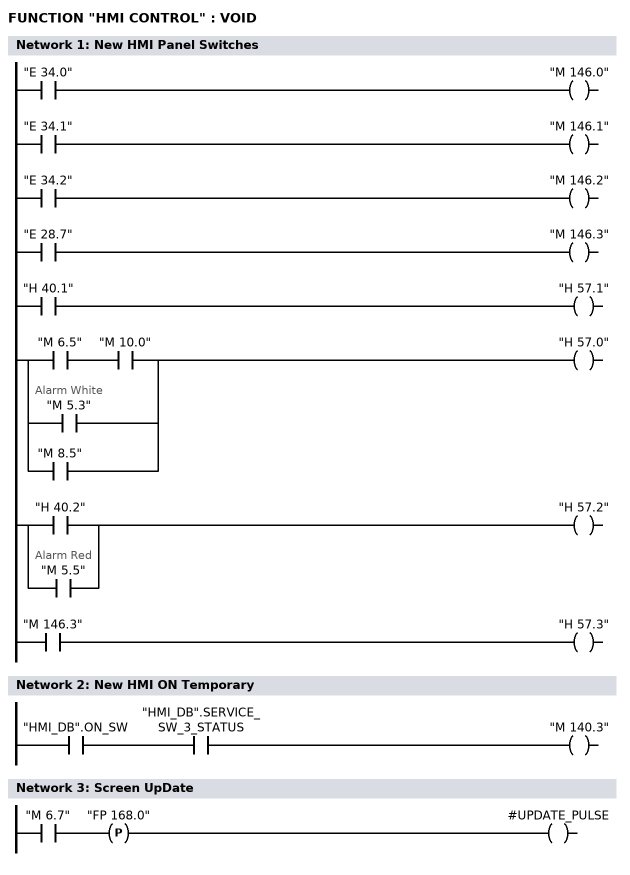

      A     "E 34.0";
      =     "M 146.0";
//;
      A     "E 34.1";
      =     "M 146.1";
//;
      A     "E 34.2";
      =     "M 146.2";
//;
      A     "E 28.7";
      =     "M 146.3";
//;
      A     "H 40.1";
      =     "H 57.1";
//;
      A(    ;
      A     "M 6.5";
      A     "M 10.0";
      )     ;
      O     "M 5.3"; // Alarm White
      O     "M 8.5";
      =     "H 57.0";
//;
      A     "H 40.2";
      O     "M 5.5"; // Alarm Red
      =     "H 57.2";
//;
      A     "M 146.3";
      =     "H 57.3";
NETWORK
TITLE =New HMI ON Temporary

      A     "HMI_DB".ON_SW;
      A     "HMI_DB".SERVICE_SW_3_STATUS;
      =     "M 140.3";
NETWORK
TITLE =Screen UpDate

      A     "M 6.7";
      FP    "FP 168.0";
      =     #UPDATE_PULSE;
NETWORK
TITLE =Screen 0 Soft Switches

      A(    ;
      L     "HMI_DB".ACTUAL_HMI_SCREEN_NO;
      L     "HMI_UPDATE".HMI_MAIN_PAGE_GRAPHIC;
      <>I   ;
      )     ;
      O     #UPDATE_PULSE;
      JNB   MAIN;
NETWORK
TITLE =Service Switch Status - Screen 0 SSW Inputs
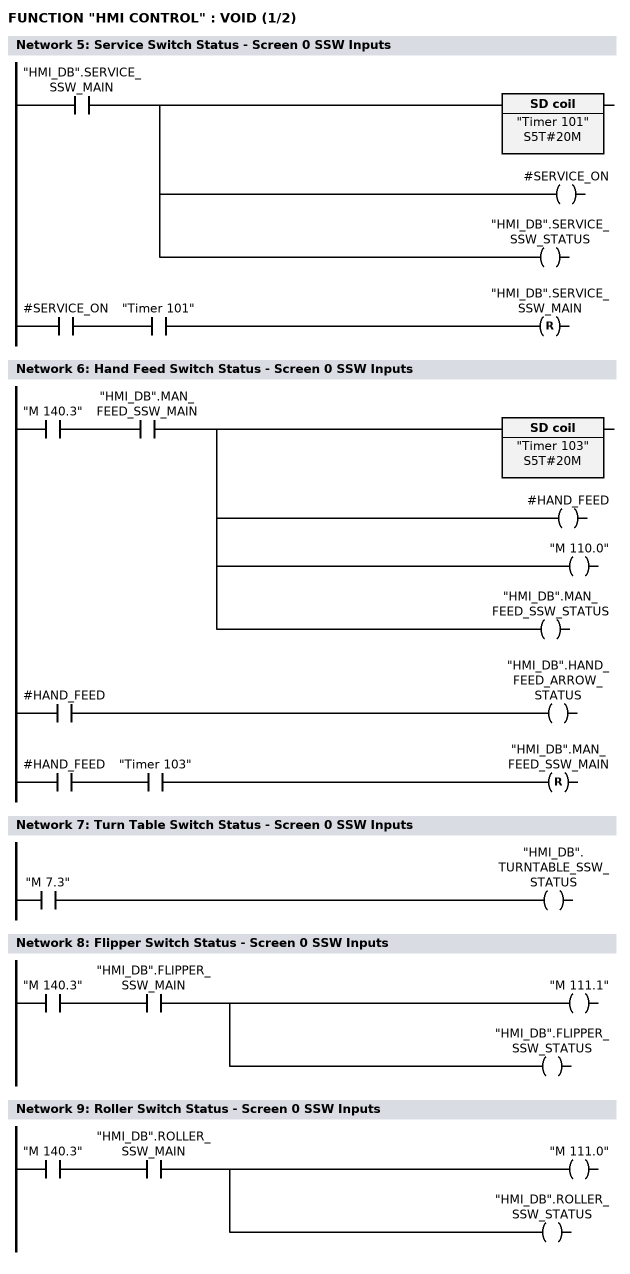

      A     "HMI_DB".SERVICE_SSW_MAIN;
      L     S5T#20M;
      SD    "Timer 101";
      =     #SERVICE_ON;
      =     "HMI_DB".SERVICE_SSW_STATUS;
//;
      A     #SERVICE_ON;
      A     "Timer 101";
      R     "HMI_DB".SERVICE_SSW_MAIN;
NETWORK
TITLE =Hand Feed Switch Status - Screen 0 SSW Inputs

      A     "M 140.3";
      A     "HMI_DB".MAN_FEED_SSW_MAIN;
      L     S5T#20M;
      SD    "Timer 103";
      =     #HAND_FEED;
      =     "M 110.0";
      =     "HMI_DB".MAN_FEED_SSW_STATUS;
//;
      A     #HAND_FEED;
      =     "HMI_DB".HAND_FEED_ARROW_STATUS;
//;
      A     #HAND_FEED;
      A     "Timer 103";
      R     "HMI_DB".MAN_FEED_SSW_MAIN;
NETWORK
TITLE =Turn Table Switch Status - Screen 0 SSW Inputs

      A     "M 7.3";
      =     "HMI_DB".TURNTABLE_SSW_STATUS;
NETWORK
TITLE =Flipper Switch Status - Screen 0 SSW Inputs

      A     "M 140.3";
      A     "HMI_DB".FLIPPER_SSW_MAIN;
      =     "M 111.1";
      =     "HMI_DB".FLIPPER_SSW_STATUS;
NETWORK
TITLE =Roller Switch Status - Screen 0 SSW Inputs

      A     "M 140.3";
      A     "HMI_DB".ROLLER_SSW_MAIN;
      =     "M 111.0";
      =     "HMI_DB".ROLLER_SSW_STATUS;
NETWORK
TITLE =HMI Service Switch Reset
//HMI Service Switch Reset when 2145 Exits Packets + 10s Delay
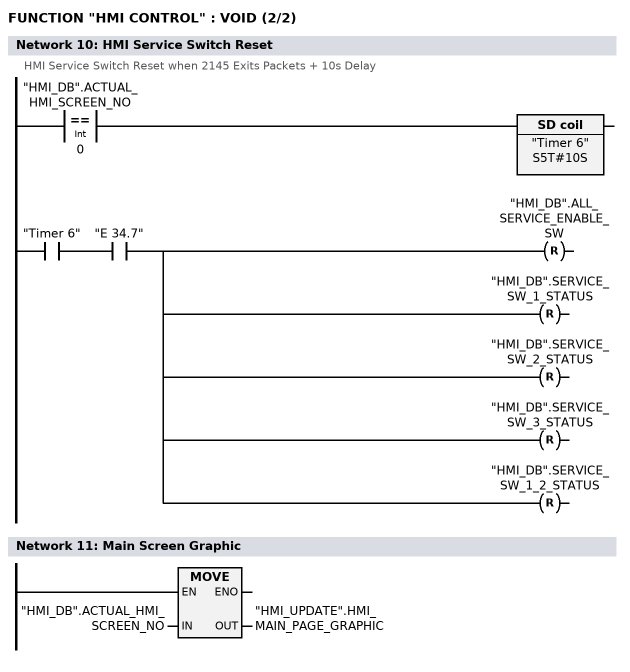
      A(    ;
      L     "HMI_DB".ACTUAL_HMI_SCREEN_NO;
      L     0;
      ==I   ;
      )     ;
      L     S5T#10S;
      SD    "Timer 6";
//;
      A     "Timer 6";
      A     "E 34.7";
      R     "HMI_DB".ALL_SERVICE_ENABLE_SW;
      R     "HMI_DB".SERVICE_SW_1_STATUS;
      R     "HMI_DB".SERVICE_SW_2_STATUS;
      R     "HMI_DB".SERVICE_SW_3_STATUS;
      R     "HMI_DB".SERVICE_SW_1_2_STATUS;
NETWORK
TITLE =Main Screen Graphic


      L     "HMI_DB".ACTUAL_HMI_SCREEN_NO;
      T     "HMI_UPDATE".HMI_MAIN_PAGE_GRAPHIC;

MAIN: NOP   0;
END_FUNCTION

FUNCTION "HMI COMMS" : VOID
TITLE =HMI Communications
//OMRON NS12  on DB12
NAME : HMI_COMM
VERSION : 0.1


VAR_TEMP
  UPDATE_PULSE_0 : BOOL ;
  UPDATE_PULSE_1 : BOOL ;
  UPDATE_PULSE_2 : BOOL ;
  UPDATE_PULSE_3 : BOOL ;
  UPDATE_PULSE_4 : BOOL ;
  UPDATE_PULSE_5 : BOOL ;
  UPDATE_PULSE_6 : BOOL ;
  UPDATE_1 : BOOL ;
  UPDATE_2 : BOOL ;
  UPDATE_3 : BOOL ;
  UPDATE_4 : BOOL ;
  UPDATE_5 : BOOL ;
  UPDATE_6 : BOOL ;
  UPDATE_7 : BOOL ;
  UPDATE_8 : BOOL ;
  UPDATE_9 : BOOL ;
  UPDATE_10 : BOOL ;
  UPDATE_11 : BOOL ;
  UPDATE_12 : BOOL ;
  UPDATE_13 : BOOL ;
  TEMP1 : BOOL ;
  TEST : BOOL ;
  CONVEYOR_0_COLOR : BYTE ;
  ELEVATOR_COLOR : BYTE ;
  CONVEYOR_1_COLOR : BYTE ;
  CONVEYOR_2_COLOR : BYTE ;
  CONVEYOR_3_COLOR : BYTE ;
  CONVEYOR_4_COLOR : BYTE ;
  CONVEYOR_5_COLOR : BYTE ;
  CONVEYOR_6_COLOR : BYTE ;
  CONVEYOR_7_COLOR : BYTE ;
  CONVEYOR_8_COLOR : BYTE ;
  CONVEYOR_9_COLOR : BYTE ;
  PUSHER_2_COLOR : BOOL ;
  CONVEYOR_11_COLOR : BYTE ;
  CONVEYOR_12_COLOR : BYTE ;
  CONVEYOR_13_COLOR : BYTE ;
  CONVEYOR_21_COLOR : BYTE ;
  CONVEYOR_22_COLOR : BYTE ;
  CONVEYOR_23_COLOR : BYTE ;
  CONVEYOR_10_COLOR : BYTE ;
  NEW_ORDER_COLOR : BYTE ;
END_VAR
BEGIN
NETWORK
TITLE =HMI - UpDate Timing
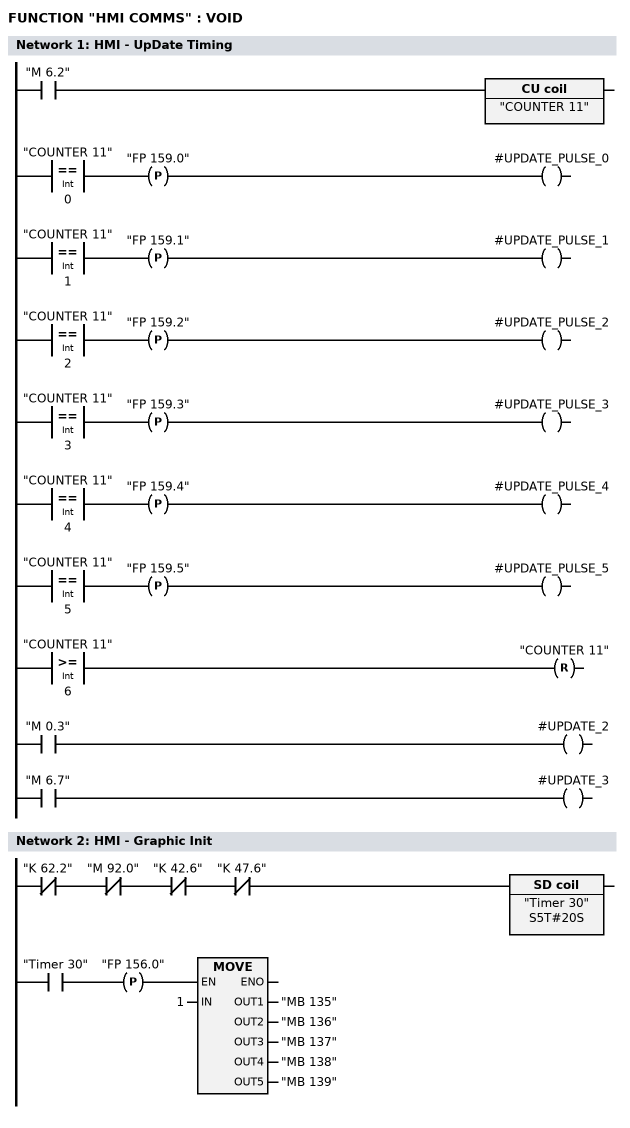

      A     "M 6.2";
      CU    "COUNTER 11";
//;
      A(    ;
      L     "COUNTER 11";
      L     0;
      ==I   ;
      )     ;
      FP    "FP 159.0";
      =     #UPDATE_PULSE_0;
//;
      A(    ;
      L     "COUNTER 11";
      L     1;
      ==I   ;
      )     ;
      FP    "FP 159.1";
      =     #UPDATE_PULSE_1;
//;
      A(    ;
      L     "COUNTER 11";
      L     2;
      ==I   ;
      )     ;
      FP    "FP 159.2";
      =     #UPDATE_PULSE_2;
//;
      A(    ;
      L     "COUNTER 11";
      L     3;
      ==I   ;
      )     ;
      FP    "FP 159.3";
      =     #UPDATE_PULSE_3;
//;
      A(    ;
      L     "COUNTER 11";
      L     4;
      ==I   ;
      )     ;
      FP    "FP 159.4";
      =     #UPDATE_PULSE_4;
//;
      A(    ;
      L     "COUNTER 11";
      L     5;
      ==I   ;
      )     ;
      FP    "FP 159.5";
      =     #UPDATE_PULSE_5;
//;
      A(    ;
      L     "COUNTER 11";
      L     6;
      >=I   ;
      )     ;
      R     "COUNTER 11";
//;;
      A     "M 0.3";
      =     #UPDATE_2;
//;
      A     "M 6.7";
      =     #UPDATE_3;
NETWORK
TITLE =HMI - Graphic Init

      AN    "K 62.2";
      AN    "M 92.0";
      AN    "K 42.6";
      AN    "K 47.6";
      L     S5T#20S;
      SD    "Timer 30";
//;
      A     "Timer 30";
      FP    "FP 156.0";
      JNB   K622;
      L     1;
      T     "MB 135";
      T     "MB 136";
      T     "MB 137";
      T     "MB 138";
      T     "MB 139";

K622: NOP   0;
NETWORK
TITLE =HMI - Doors Monitor

      ON    "E 4.6";
      ON    "E 9.0";
      ON    "E 12.5";
      O     #UPDATE_PULSE_0;
      JNB   DOOR;
      AN    "E 4.6";
      =     "HMI_DB".ELEVATOR_DOOR_STATUS;
//;
      AN    "E 9.0";
      =     "HMI_DB".FLIPPER_DOOR_STATUS;
//;
      AN    "E 12.5";
      =     "HMI_DB".LOADER_DOOR_STATUS;

DOOR: NOP   0;
NETWORK
TITLE =HMI - E-Stop Monitor

      O     "M 1.0";
      O     "M 1.1";
      O     "M 1.2";
      O     "M 1.3";
      O     #UPDATE_PULSE_1;
      JNB   ESTP;
      A     "M 1.0";
      =     "HMI_DB".E_STOP_CONSOLE_STATUS;
//;
      A     "M 1.1";
      =     "HMI_DB".E_STOP_LOADER_STATUS;
//;
      A     "M 1.2";
      =     "HMI_DB".E_STOP_ELEVATOR_STATUS;
//;
      A     "M 1.3";
      =     "HMI_DB".E_STOP_FLIPPER_STATUS;

ESTP: NOP   0;
NETWORK
TITLE =HMI - Motors Fault Status

      A(    ;
      L     "MW 2";
      L     0;
      <>I   ;
      O     ;
      L     "MB 4";
      L     0;
      <>I   ;
      )     ;
      O     "M 7.0";
      O     "M 7.1";
      O     "M 7.2";
      O     #UPDATE_PULSE_2;
      JNB   MTRF;
      A     "M 2.0";
      =     "HMI_DB".CONVEYOR_0_MOTOR_STATUS;
//;
      A     "M 2.1";
      =     "HMI_DB".PUSHER_0_MOTOR_STATUS;
//;
      A     "M 2.2";
      =     "HMI_DB".ELEVATOR_MOTOR_STATUS;
//;
      A     "M 2.3";
      =     "HMI_DB".PUSHER_1_MOTOR_STATUS;
//;
      A     "M 2.4";
      =     "HMI_DB".CONVEYOR_1_MOTOR_STATUS;
//;
      A     "M 2.5";
      =     "HMI_DB".CONVEYOR_2B_MOTOR_STATUS;
//;
      A     "M 2.6";
      =     "HMI_DB".CONVEYOR_2R_MOTOR_STATUS;
//;
      A     "M 2.7";
      =     "HMI_DB".CONVEYOR_3_MOTOR_STATUS;
//;
      A     "M 3.0";
      =     "HMI_DB".CONVEYOR_4_MOTOR_STATUS;
//;
      A     "M 3.1";
      =     "HMI_DB".CONVEYOR_5_MOTOR_STATUS;
//;
      A     "M 3.2";
      =     "HMI_DB".CONVEYOR_6_MOTOR_STATUS;
//;
      A     "M 3.3";
      =     "HMI_DB".CONVEYOR_7_MOTOR_STATUS;
//;
      A     "M 3.4";
      =     "HMI_DB".FLIPPER_MOTOR_STATUS;
//;
      A     "M 3.5";
      =     "HMI_DB".CONVEYOR_8_MOTOR_STATUS;
//;
      A     "M 3.6";
      =     "HMI_DB".TURNTABLE_MOTOR_STATUS;
//;
      A     "M 3.7";
      =     "HMI_DB".CONVEYOR_9_MOTOR_STATUS;
//;
      A     "M 4.0";
      =     "HMI_DB".PUSHER_2_MOTOR_STATUS;
//;
      A     "M 4.1";
      =     "HMI_DB".CONVEYOR_10_MOTOR_STATUS;
//;
      A     "M 4.2";
      =     "HMI_DB".CONVEYOR_11_MOTOR_STATUS;
//;
      A     "M 4.3";
      =     "HMI_DB".CONVEYOR_12_MOTOR_STATUS;
//;
      A     "M 4.4";
      =     "HMI_DB".CONVEYOR_13_MOTOR_STATUS;
//;
      A     "M 4.5";
      =     "HMI_DB".CONVEYOR_21_MOTOR_STATUS;
//;
      A     "M 4.6";
      =     "HMI_DB".CONVEYOR_22_MOTOR_STATUS;
//;
      A     "M 4.7";
      =     "HMI_DB".CONVEYOR_23_MOTOR_STATUS;
//;
      A     "M 7.0";
      =     "HMI_DB".LOADER_LIFT_MOTOR_STATUS;
//;
      A     "M 7.1";
      =     "HMI_DB".LOADER_FING_MOTOR_STATUS;
//;
      A     "M 7.2";
      =     "HMI_DB".LOADER_BELT_MOTOR_STATUS;

MTRF: NOP   0;
NETWORK
TITLE =HMI Light Barriers Status - Conveyors 1, 2, 3 LBs

      A(    ;
      L     IW     5;
      L     "HMI_UPDATE".HMI_GRAPHIC_TOTAL_1;
      <>I   ;
      O     #UPDATE_PULSE_3;
      )     ;
      JNB   LBS1;
      A     "B 5.4";
      =     "HMI_DB".LIGHT_BARRIER_1_STATUS;
//;
      A     "B 5.5";
      =     "HMI_DB".LIGHT_BARRIER_2_STATUS;
//;
      A     "B 6.0";
      =     "HMI_DB".LIGHT_BARRIER_3_STATUS;
//;
      A     "B 6.1";
      =     "HMI_DB".LIGHT_BARRIER_4_STATUS;
//;
      A     "B 6.2";
      =     "HMI_DB".LIGHT_BARRIER_5_STATUS;
//;
      A     "B 6.4";
      =     "HMI_DB".LIGHT_BARRIER_6_STATUS;
//;
      A     "B 5.2";
      =     "HMI_DB".LIGHT_BARRIER_B_STATUS;
//;
      A     "B 5.1";
      =     "HMI_DB".LIGHT_BARRIER_A_STATUS;
//;
      L     IW     5;
      T     "HMI_UPDATE".HMI_GRAPHIC_TOTAL_1;

LBS1: NOP   0;
NETWORK
TITLE =HMI Light Barriers Status - Conveyors 4, 5, 6, 7, 8, 9 LBs

      A(    ;
      L     IW     6;
      L     "HMI_UPDATE".HMI_GRAPHIC_TOTAL_2;
      <>I   ;
      O     #UPDATE_PULSE_4;
      )     ;
      O     "B 8.2";
      JNB   LBS2;
      A     "B 6.7";
      =     "HMI_DB".LIGHT_BARRIER_7_STATUS;
//;
      A     "B 7.0";
      =     "HMI_DB".LIGHT_BARRIER_8_STATUS;
//;
      A     "B 7.1";
      =     "HMI_DB".LIGHT_BARRIER_9_STATUS;
//;
      A     "B 7.2";
      =     "HMI_DB".LIGHT_BARRIER_10_STATUS;
//;
      A     "B 7.3";
      =     "HMI_DB".LIGHT_BARRIER_11_STATUS;
//;
      A     "B 7.4";
      =     "HMI_DB".LIGHT_BARRIER_12_STATUS;
//;
      A     "B 8.2";
      =     "HMI_DB".LIGHT_BARRIER_13_STATUS;
//;
      L     IW     6;
      T     "HMI_UPDATE".HMI_GRAPHIC_TOTAL_2;

LBS2: NOP   0;
NETWORK
TITLE =HMI Light Barriers Status - Conveyors 10, 11, 12, 13, 21, 22, 23

      A(    ;
      L     IW     9;
      L     IW    12;
      +I    ;
      L     IB    15;
      +I    ;
      L     "HMI_UPDATE".HMI_FEED_GRAPHIC;
      <>I   ;
      O     #UPDATE_PULSE_5;
      )     ;
      JNB   LBS3;
      A     "B 9.6";
      =     "HMI_DB".LIGHT_BARRIER_14_STATUS;
//;
      A     "B 9.7";
      =     "HMI_DB".LIGHT_BARRIER_15_STATUS;
//;
      A     "B 10.3";
      =     "HMI_DB".LIGHT_BARRIER_16_STATUS;
//;
      A     "B 10.4";
      =     "HMI_DB".LIGHT_BARRIER_17_STATUS;
//;
      A     "B 10.5";
      =     "HMI_DB".LIGHT_BARRIER_18_STATUS;
//;
      A     "B 10.6";
      =     "HMI_DB".LIGHT_BARRIER_19_STATUS;
//;
      A     "B 10.7";
      =     "HMI_DB".LIGHT_BARRIER_20_STATUS;
//;
      A     "B 11.0";
      =     "HMI_DB".LIGHT_BARRIER_21_STATUS;
//;
      A     "B 11.1";
      =     "HMI_DB".LIGHT_BARRIER_22_STATUS;
//;
      A     "B 11.2";
      =     "HMI_DB".LIGHT_BARRIER_23_STATUS;
//;
      A     "B 12.3";
      =     "HMI_DB".LIGHT_BARRIER_24_STATUS;
//;
      A     "B 13.0";
      =     "HMI_DB".LIGHT_BARRIER_25_STATUS;
//;
      A     "B 15.4";
      =     "HMI_DB".LIGHT_BARRIER_26_STATUS;
//;
      A     "B 15.5";
      =     "HMI_DB".LIGHT_BARRIER_27_STATUS;
//;
      A     "B 15.6";
      =     "HMI_DB".LIGHT_BARRIER_28_STATUS;
//;
      A     "B 15.7";
      =     "HMI_DB".LIGHT_BARRIER_29_STATUS;
//;
      L     IW     9;
      L     IW    12;
      +I    ;
      L     IB    15;
      +I    ;
      T     "HMI_UPDATE".HMI_FEED_GRAPHIC;

LBS3: NOP   0;
NETWORK
TITLE =HMI Light Barriers Status - Conveyors 0 LBs

      A(    ;
      L     QB    62;
      L     "HMI_UPDATE".HMI_MOTOR_TOTAL_1;
      <>I   ;
      O     #UPDATE_PULSE_0;
      )     ;
      O     "B 8.2";
      JNB   LBS4;
      A     "E 34.7";
      =     "HMI_DB".PACKETIZER_GATE_STATUS;
//;
      A     "B 35.2";
      =     "HMI_DB".LIGHT_BARRIER_30_STATUS;
//;
      A     "B 35.3";
      =     "HMI_DB".LIGHT_BARRIER_31_STATUS;
//;
      A     "B 35.4";
      =     "HMI_DB".LIGHT_BARRIER_32_STATUS;
//;
      L     QB    62;
      T     "HMI_UPDATE".HMI_MOTOR_TOTAL_1;

LBS4: NOP   0;
NETWORK
TITLE =HMI Prox Sensors Status - Elevator - Proxs

      A(    ;
      L     IB     4;
      L     "HMI_UPDATE".HMI_ELEVATOR_PROXS;
      <>I   ;
      O     #UPDATE_PULSE_1;
      )     ;
      JNB   PRX1;
      AN    "P 4.0";
      =     "HMI_DB".PROX_1_STATUS;
//;
      AN    "P 4.1";
      =     "HMI_DB".PROX_2_STATUS;
//;
      AN    "P 4.2";
      =     "HMI_DB".PROX_3_STATUS;
//;
      AN    "P 4.3";
      =     "HMI_DB".PROX_4_STATUS;
//;
      AN    "P 4.4";
      =     "HMI_DB".PROX_5_STATUS;
//;
      AN    "P 4.5";
      =     "HMI_DB".PROX_6_STATUS;
//;
      L     IB     4;
      T     "HMI_UPDATE".HMI_ELEVATOR_PROXS;

PRX1: NOP   0;
NETWORK
TITLE =HMI Prox Sensors Status - Flipper / TurnTable - Proxs

      A(    ;
      L     IW     8;
      L     "HMI_UPDATE".HMI_FLIPPER_PROXS;
      <>I   ;
      O     #UPDATE_PULSE_2;
      )     ;
      JNB   PRX2;
      AN    "P 8.0";
      =     "HMI_DB".PROX_8_STATUS;
//;
      AN    "P 8.1";
      =     "HMI_DB".PROX_7_STATUS;
//;
      AN    "P 8.5";
      =     "HMI_DB".PROX_9_STATUS;
//;
      AN    "P 8.6";
      =     "HMI_DB".PROX_10_STATUS;
//;
      AN    "P 9.2";
      =     "HMI_DB".PROX_11_STATUS;
//;
      AN    "P 9.3";
      =     "HMI_DB".PROX_12_STATUS;
//;
      L     IW     8;
      T     "HMI_UPDATE".HMI_FLIPPER_PROXS;

PRX2: NOP   0;
NETWORK
TITLE =HMI Prox Sensors Status - Pusher 2 / Pivot 10 - Proxs

      A(    ;
      L     IB    10;
      L     IB    15;
      +I    ;
      L     "HMI_UPDATE".HMI_PUSHER_PROXS;
      <>I   ;
      O     #UPDATE_PULSE_3;
      )     ;
      JNB   PRX3;
      AN    "P 10.0";
      =     "HMI_DB".PROX_13_STATUS;
//;
      AN    "P 10.1";
      =     "HMI_DB".PROX_14_STATUS;
//;
      A     "P 15.0";
      =     "HMI_DB".PROX_15_STATUS;
//;
      A     "P 15.1";
      =     "HMI_DB".PROX_16_STATUS;
//;
      L     IB    10;
      L     IB    15;
      +I    ;
      T     "HMI_UPDATE".HMI_PUSHER_PROXS;

PRX3: NOP   0;
NETWORK
TITLE =HMI Prox Sensors Status - Feeder - Proxs

      A(    ;
      L     IW    11;
      L     IB    13;
      +I    ;
      L     "HMI_UPDATE".HMI_FEEDER_PROXS;
      <>I   ;
      O     #UPDATE_PULSE_4;
      )     ;
      JNB   PRX4;
      AN    "P 13.2";
      =     "HMI_DB".PROX_17_STATUS;
//;
      AN    "P 13.1";
      =     "HMI_DB".PROX_18_STATUS;
//;
      AN    "P 11.4";
      =     "HMI_DB".PROX_19_STATUS;
//;
      AN    "P 11.5";
      =     "HMI_DB".PROX_20_STATUS;
//;
      AN    "P 11.6";
      =     "HMI_DB".PROX_21_STATUS;
//;
      AN    "P 11.7";
      =     "HMI_DB".PROX_22_STATUS;
//;
      A     "P 12.0";
      =     "HMI_DB".PROX_23_STATUS;
//;
      A     "P 12.1";
      =     "HMI_DB".PROX_24_STATUS;
//;
      L     IW    11;
      L     IB    13;
      +I    ;
      T     "HMI_UPDATE".HMI_FEEDER_PROXS;

PRX4: NOP   0;
NETWORK
TITLE =HMI - Pusher 0 - Graphic

      A(    ;
      O     "K 62.2";
      O     "K 62.3";
      O     #UPDATE_PULSE_5;
      )     ;
      JNB   PUS0;
      A     "K 62.2";
      AN    "K 62.3";
      A     "M 6.1";
      AN(   ;
      L     "MB 135";
      L     L#128;
      >=I   ;
      )     ;
      FP    "FP 156.1";
      JNB   E622;
      L     "MB 135";
      SLW   1;
      T     "MB 135";

E622: NOP   0;

      A     "K 62.3";
      AN    "K 62.2";
      A     "M 6.1";
      AN(   ;
      L     "MB 135";
      L     L#1;
      <=I   ;
      )     ;
      FP    "FP 156.2";
      JNB   R623;
      L     "MB 135";
      SRW   1;
      T     "MB 135";

R623: NOP   0;

      A     "M 6.1";
      FP    "HMI_DB".FP133;
      JNB   P133;
      L     L#255;
      L     "MB 135";
      -I    ;
      T     DB12.DBB    4;

P133: NOP   0;

PUS0: NOP   0;
NETWORK
TITLE =HMI - Elevator - Graphic

      A(    ;
      O     "M 92.0";
      O     "M 92.1";
      O     #UPDATE_PULSE_0;
      )     ;
      JNB   ELEV;
      A     "M 92.0";
      AN    "M 92.1";
      A     "M 6.2";
      AN(   ;
      L     "MB 136";
      L     L#128;
      >=I   ;
      )     ;
      FP    "FP 156.3";
      JNB   R420;
      L     "MB 136";
      SLW   1;
      T     "MB 136";

R420: NOP   0;

      A     "M 92.1";
      AN    "M 92.0";
      A     "M 6.2";
      AN(   ;
      L     "MB 136";
      L     L#1;
      <=I   ;
      )     ;
      FP    "FP 156.4";
      JNB   F420;
      L     "MB 136";
      SRW   1;
      T     "MB 136";

F420: NOP   0;

      A     "M 6.2";
      FP    "HMI_DB".FP134;
      JNB   P134;
      L     L#255;
      L     "MB 136";
      -I    ;
      T     DB12.DBB    5;

P134: NOP   0;

ELEV: NOP   0;
NETWORK
TITLE =HMI - Pusher 1 - Graphic

      A(    ;
      O     "K 42.6";
      O     "K 42.7";
      O     #UPDATE_PULSE_1;
      )     ;
      JNB   PUS1;
      A     "K 42.6";
      AN    "K 42.7";
      A     "M 6.1";
      AN(   ;
      L     "MB 137";
      L     L#128;
      >=I   ;
      )     ;
      FP    "FP 156.5";
      JNB   E426;
      L     "MB 137";
      SLW   1;
      T     "MB 137";

E426: NOP   0;

      A     "K 42.7";
      AN    "K 42.6";
      A     "M 6.1";
      AN(   ;
      L     "MB 137";
      L     L#1;
      <=I   ;
      )     ;
      FP    "FP 156.6";
      JNB   R427;
      L     "MB 137";
      SRW   1;
      T     "MB 137";

R427: NOP   0;

      A     "M 6.1";
      FP    "HMI_DB".FP135;
      JNB   P135;
      L     L#255;
      L     "MB 137";
      -I    ;
      T     DB12.DBB    6;

P135: NOP   0;

PUS1: NOP   0;
NETWORK
TITLE =HMI - Flipper Graphic

      A(    ;
      O     "K 46.0";
      O     "K 46.1";
      O     #UPDATE_PULSE_2;
      )     ;
      JNB   FLPN;
      L     3;
      A     "P 8.0";
      A     "P 8.1";
      JC    FLIP;
      L     0;

FLIP: T     "HMI_DB".FLIPPER_TURN_COLOR;

      L     1;
      AN    "P 8.0";
      A     "P 8.1";
      JC    CCW1;
      L     "HMI_DB".FLIPPER_TURN_COLOR;

CCW1: T     "HMI_DB".FLIPPER_CCW;

      L     1;
      AN    "P 8.1";
      A     "P 8.0";
      JC    CW1;
      L     "HMI_DB".FLIPPER_TURN_COLOR;

CW1:  T     "HMI_DB".FLIPPER_CW;

      L     6;
      A     "M 42.0";
      JC    FLON;
      L     9;

FLON: T     "HMI_DB".FLIPPER_COLOR;

FLPN: NOP   0;
NETWORK
TITLE =HMI - TurnTable Graphic

      A(    ;
      O     "A 47.0";
      O     "A 47.1";
      O     #UPDATE_PULSE_3;
      )     ;
      JNB   TURN;
      A(    ;
      ON    "P 9.2";
      ON    "P 9.3";
      )     ;
      S     "HMI_DB".TURNTABLE_DELIV_POSITION;
//;
      A(    ;
      ON    "P 8.5";
      ON    "P 8.6";
      )     ;
      R     "HMI_DB".TURNTABLE_DELIV_POSITION;
//;
      AN    "M 7.3";
      =     "HMI_DB".TURNTABLE_REVERSE_ARROW;
//;
      A     "M 7.3";
      =     "HMI_DB".TURNTABLE_DIR_SELECT_SW;

TURN: NOP   0;

NETWORK
TITLE =HMI - Pusher 2 - Graphic

      A(    ;
      O     "K 47.6";
      O     "K 47.7";
      O     #UPDATE_PULSE_4;
      )     ;
      JNB   PUS2;
      A     "K 47.6";
      AN    "K 47.7";
      A     "M 6.1";
      AN(   ;
      L     "MB 138";
      L     L#128;
      >=I   ;
      )     ;
      FP    "FP 156.7";
      JNB   E476;
      L     "MB 138";
      SLW   1;
      T     "MB 138";

E476: NOP   0;

      A     "K 47.7";
      AN    "K 47.6";
      A     "M 6.1";
      AN(   ;
      L     "MB 138";
      L     L#1;
      <=I   ;
      )     ;
      FP    "FP 157.0";
      JNB   R477;
      L     "MB 138";
      SRW   1;
      T     "MB 138";

R477: NOP   0;

      A     "M 6.1";
      FP    "HMI_DB".FP140;
      JNB   P140;
      L     L#255;
      L     "MB 138";
      -I    ;
      T     DB12.DBB    7;

P140: NOP   0;

PUS2: NOP   0;
NETWORK
TITLE =HMI - Pivot Graphic

      A(    ;
      O     "K 53.0";
      O     "K 53.1";
      O     #UPDATE_PULSE_5;
      )     ;
      JNB   PIVO;
      AN    "P 15.1";
      =     DB12.DBX   88.1;
//;
      AN    "P 15.0";
      =     DB12.DBX   88.0;
//;
      AN    "P 15.0";
      AN    "P 15.1";
      =     DB12.DBX   88.2;

PIVO: NOP   0;
NETWORK
TITLE =HMI - Feeder Graphic

      A(    ;
      L     IW    11;
      L     IB    13;
      +I    ;
      L     "HMI_UPDATE".HMI_FEEDER_GRAPHIC;
      <>I   ;
      O     #UPDATE_PULSE_0;
      )     ;
      JNB   FEED;

      A     "P 13.2";
      AN    "P 11.4";
      O     ;
      A     "P 11.5";
      AN    "P 11.4";
      JNB   M131;
      L     L#64;
      T     "MB 139";

M131: NOP   0;

      AN    "P 13.2";
      AN    "P 13.1";
      AN    "P 11.4";
      JNB   M132;
      L     L#128;
      T     "MB 139";

M132: NOP   0;

      AN    "P 11.4";
      AN    "P 11.5";
      JNB   M114;
      L     L#32;
      T     "MB 139";

M114: NOP   0;

      A     "P 11.4";
      AN    "P 11.5";
      A     "A 50.1";
      S     "M 70.5";
//;
      A(    ;
      A     "M 70.6";
      A     "A 50.0";
      AN    "P 11.5";
      O     ;
      A     "M 70.5";
      A     "A 50.1";
      )     ;
      JNB   M115;
      L     L#16;
      T     "MB 139";
      R     "M 70.6";

M115: NOP   0;

      A     "P 11.7";
      AN    "P 11.6";
      A     "A 50.0";
      S     "M 70.6";
//;
      A(    ;
      A     "M 70.5";
      A     "A 50.1";
      AN    "P 11.6";
      O     ;
      A     "M 70.6";
      A     "A 50.0";
      )     ;
      JNB   M116;
      L     L#8;
      T     "MB 139";
      R     "M 70.5";

M116: NOP   0;

      AN    "E 12.2";
      AN    "P 11.7";
      AN    "P 12.1";
      JNB   M117;
      L     L#4;
      T     "MB 139";

M117: NOP   0;

      AN    "E 12.2";
      AN    "P 11.7";
      A     "P 12.1";
      JNB   M121;
      L     L#6;
      T     "MB 139";

M121: NOP   0;

      A     "E 12.2";
      AN    "P 11.7";
      A     "P 12.1";
      JNB   M122;
      L     L#1;
      T     "MB 139";

M122: NOP   0;

      A     "M 6.2";
      FP    "HMI_DB".FP141;
      JNB   P141;
      L     L#255;
      L     "MB 139";
      -I    ;
      T     DB12.DBB   19;

P141: NOP   0;

      L     IW    11;
      L     IB    13;
      +I    ;
      T     "HMI_UPDATE".HMI_FEEDER_GRAPHIC;

FEED: NOP   0;
NETWORK
TITLE =HMI - Motor Run Status

      A(    ;
      L     QW    42;
      L     QW    44;
      +I    ;
      L     QW    46;
      +I    ;
      L     QW    48;
      +I    ;
      L     QW    50;
      +I    ;
      L     QB    53;
      +I    ;
      L     QB    54;
      +I    ;
      L     "HMI_UPDATE".HMI_MOTOR_GRAPHIC;
      <>I   ;
      O     #UPDATE_PULSE_1;
      )     ;
      JNB   MTR;
      O     "K 62.0";
      O     "K 62.1";
      L     0;
      JCN   K620;
      A     "K 62.0";
      L     3;
      JC    K620;
      L     6;
K620: T     "HMI_DB".CONV_0_COLOR_WORD;

      L     5;
      A     "M 14.7";
      O     "M 100.2";
      JC    E00;
      L     0;
E00:  T     #ELEVATOR_COLOR;

      L     #ELEVATOR_COLOR;
      O     "M 92.0";
      O     "M 92.1";
      JCN   Q420;
      A     "M 92.0";
      L     3;
      JC    Q420;
      L     6;
Q420: T     "HMI_DB".ELEVATOR_COLOR_WORD;

      L     0;
      A(    ;
      O     "K 42.6";
      O     "K 42.7";
      )     ;
      JCN   Q427;
      L     3;
Q427: T     "HMI_DB".PUSHER_1_COLOR_WORD;

      L     0;
      A     "A 43.0";
      JCN   Q430;
      L     3;
Q430: T     "HMI_DB".CONV_1_COLOR_WORD;

      L     5;
      A     "M 22.7";
      O     "M 100.5";
      JC    C02;
      L     0;
C02:  T     #CONVEYOR_2_COLOR;

      L     #CONVEYOR_2_COLOR;
      A     "K 43.4";
      JCN   Q434;
      L     3;
Q434: T     "HMI_DB".CONV_2_BELT_COLOR_WORD;

      L     0;
      A     "Y 43.6";
      JCN   Q436;
      L     3;
Q436: T     "HMI_DB".LIFT_ROLLER_2_COLOR_WORD;

      L     0;
      A     "K 43.5";
      JCN   Q435;
      L     3;
Q435: T     "HMI_DB".CONV_2_ROLLER_COLOR_WORD;

      L     0;
      A     "A 44.0";
      JCN   Q440;
      L     3;
Q440: T     "HMI_DB".CONV_3_COLOR_WORD;

      L     5;
      A     "M 30.7";
      O     "M 102.0";
      JC    C04;
      L     0;
C04:  T     #CONVEYOR_4_COLOR;

      L     #CONVEYOR_4_COLOR;
      A     "A 44.3";
      AN    "M 31.5";
      JCN   Q443;
      L     6;
Q443: T     "HMI_DB".CONV_4_COLOR_WORD;

      A     "A 44.3";
      A     "M 31.5";
      JNB   M315;
      L     3;
      T     "HMI_DB".CONV_4_COLOR_WORD;

M315: NOP   0;

      L     0;
      A     "A 45.0";
      JCN   Q450;
      L     3;
Q450: T     "HMI_DB".CONV_5_COLOR_WORD;

      L     5;
      A     "M 38.7";
      O     "M 102.2";
      JC    C06;
      L     0;
C06:  T     #CONVEYOR_6_COLOR;

      L     #CONVEYOR_6_COLOR;
      A     "A 45.3";
      JCN   Q453;
      L     3;
Q453: T     "HMI_DB".CONV_6_COLOR_WORD;

      L     5;
      A     "M 42.7";
      O     "M 102.3";
      JC    C07;
      L     0;
C07:  T     #CONVEYOR_7_COLOR;

      L     #CONVEYOR_7_COLOR;
      A     "A 45.6";
      JCN   Q456;
      L     3;
Q456: T     "HMI_DB".CONV_7_COLOR_WORD;

      L     0;
      A(    ;
      O     "K 46.0";
      O     "K 46.1";
      )     ;
      JCN   Q461;
      L     3;
Q461: T     "HMI_DB".FLIPPER_COLOR_WORD;

      L     0;
      A(    ;
      O     "A 47.0";
      O     "A 47.1";
      )     ;
      JCN   A470;
      L     7;

A470: T     "HMI_DB".TURN_COLOR;

//      L     0
//      AN    "M 6.2"
//      A(
//      O     "A 47.0"
//      O     "A 47.1"
//      )
//      JCN   A471
//      L     7

//A471: T     "HMI_DB".HMI_TURN_COLOR

      L     "HMI_DB".TURN_COLOR;
      A(    ;
      O     "A 46.4";
      O     "A 46.5";
      )     ;
      JCN   Q464;
      L     3;
Q464: T     "HMI_DB".CONV_8_COLOR_WORD;

      L     0;
      A     "A 47.0";
      JCN   Q470;
      L     3;
Q470: T     "HMI_DB".TURN_TABLE_COLOR_WORD;

      L     0;
      A     "K 47.5";
      JCN   Q475;
      L     3;
Q475: T     "HMI_DB".CONV_9_COLOR_WORD;

      L     0;
      A(    ;
      O     "K 47.6";
      O     "K 47.7";
      )     ;
      JCN   Q477;
      L     3;
Q477: T     "HMI_DB".PUSHER_2_COLOR_WORD;

      L     5;
      A     "M 98.1";
      O     "M 98.2";
      O     "M 106.1";
      JC    C10;
//;
      L     4;
      A     "M 55.4";
      A     "M 8.4";
      A     "M 6.5";
      JC    C10;
      L     0;

C10:  T     #CONVEYOR_10_COLOR;

      L     #CONVEYOR_10_COLOR;
      A     "A 48.0";
      A(    ;
      ON    "M 55.5";
      ON    "M 10.0";
      )     ;
      JCN   Q480;
      L     6;
Q480: T     "HMI_DB".CONV_10_COLOR_WORD;

      A     "A 48.0";
      A(    ;
      O     "M 55.5";
      O     "M 10.0";
      )     ;
      JNB   M555;
      L     3;
      T     "HMI_DB".CONV_10_COLOR_WORD;

M555: NOP   0;


      L     0;
      A     "A 48.3";
      JCN   Q483;
      L     3;
Q483: T     "HMI_DB".CONV_11_COLOR_WORD;

      L     0;
      A     "A 48.6";
      JCN   Q486;
      L     3;
Q486: T     "HMI_DB".CONV_12_COLOR_WORD;

      L     5;
      A     "M 66.7";
      O     "M 106.4";
      JC    C13;
      L     0;
C13:  T     #CONVEYOR_13_COLOR;

      L     #CONVEYOR_13_COLOR;
      A     "A 49.0";
      JCN   Q490;
      L     3;
Q490: T     "HMI_DB".CONV_13_COLOR_WORD;

      L     0;
      A     "A 53.4";
      JCN   Q534;
      L     3;
Q534: T     "HMI_DB".CONV_21_COLOR_WORD;

      L     0;
      A     "A 53.6";
      JCN   Q536;
      L     3;
Q536: T     "HMI_DB".CONV_22_COLOR_WORD;

      L     5;
      A     "M 86.7";
      O     "M 106.7";
      JC    C23;
      L     0;
C23:  T     #CONVEYOR_23_COLOR;

      L     #CONVEYOR_23_COLOR;
      A     "A 54.0";
      JCN   Q540;
      L     3;
Q540: T     "HMI_DB".CONV_23_COLOR_WORD;

      A     "M 0.7";
      =     "HMI_DB".COMPRESSED_AIR;
//;
      O     "A 50.0";
      O     "A 50.1";
      L     0;
      JCN   Q500;
      A     "A 50.0";
      L     3;
      JC    Q500;
      L     6;
Q500: T     "HMI_DB".LOADER_LIFT_COLOR_WORD;

      L     0;
      A     "A 51.0";
      JCN   Q510;
      L     3;
Q510: T     "HMI_DB".FINGERS_BELT_COLOR_WORD;

      L     QW    42;
      L     QW    44;
      +I    ;
      L     QW    46;
      +I    ;
      L     QW    48;
      +I    ;
      L     QW    50;
      +I    ;
      L     QB    53;
      +I    ;
      L     QB    54;
      +I    ;
      T     "HMI_UPDATE".HMI_MOTOR_GRAPHIC;

MTR:  NOP   0;
END_FUNCTION

FUNCTION "HMI PACKET COUNTER  NEW" : VOID
TITLE =HMI Conveyors Display Packet Counter  FC1208
//Counts are kept in "HMI_DB" (read by HMI, LIGHT BAR, C5 Re-Sync)
//Bit_0 = InFeed  /  Bit_1 = RAW Exit Sensor  /
//Transfer_Start = Transfer Step Active.
VERSION : 0.3


VAR_TEMP
  ERROR : BOOL ;
  BIT0 : BOOL ;	//Count UP Input
  XFER : BOOL ;	//Transfer Active
  DIM_31 : INT ;	//C10 Width @ 31.0 m/min [mS]
  DIM_237 : INT ;	//C10 Width @ 23.7 m/min [mS]
END_VAR
BEGIN
NETWORK
TITLE =Packet Length mm - To Conveyor 4 HMI (as FC1206)

      L     "COLLATORS DB".PacketLength_C4;
      ITD   ;
      DTR   ;
      L     6.673000e+00;
      *R    ;
      RND   ;
      T     "MW 202";
NETWORK
TITLE =C10 Packet Width [mS] - Scaled to Link & Delivery Speeds

      L     "COLLATORS DB".Packet_Width_C10_mS; // Measured @ 27.0 m/min
      L     L#27;
      *D    ;
      L     L#31;
      /D    ;
      T     #DIM_31; // @ 31.0 m/min
      L     "COLLATORS DB".Packet_Width_C10_mS;
      L     L#270;
      *D    ;
      L     L#237;
      /D    ;
      T     #DIM_237; // @ 23.7 m/min
NETWORK
TITLE =Packet Counter - Slat Conveyor 3

      A     "A 44.0";
      L     S5T#1S;
      SF    T    118; // Call Hold 1s
      A     T    118;
      JNB   M440;
      L     "HMI_DB".CONVEYOR_MAXCOUNT_L;
      T     "DEBOUNCER COUNTER DB".Conveyor_C3_Slat.Maximum_Count;
      A     "B 6.2";
      =     #BIT0;
      A     "A 44.0";
      =     #XFER;
      CALL "DE-BOUNCER / COUNTER" (
           Bit_0                    := #BIT0,
           Bit_1                    := "B 6.4",
           Transfer_Start           := #XFER,
           Error_Reset              := "M 9.1",
           Space_DX_mS              := 600,
           ReSample_DX              := 85,
           Conveyor_Type            := 1,
           Preset_MIN_mS            := 500,
           LowSpd_Dimension_mS      := 0,
           HighSpd_Dimension_mS     := 0,
           Plc_Scan_mS              := "DB UTILITY".Scan_Cycle_Previous,
           Q_Error                  := #ERROR,
           Word_Count               := "HMI_DB".CONV_3_COUNT,
           IO_DB                    := "DEBOUNCER COUNTER DB".Conveyor_C3_Slat);
M440: NOP   0;
NETWORK
TITLE =Packet Counter - Collator Conveyor 4

      A     "A 44.3";
      L     S5T#1S;
      SF    T    119; // Call Hold 1s
      A     T    119;
      JNB   M443;
      L     "HMI_DB".CONVEYOR_MAXCOUNT_L;
      T     "DEBOUNCER COUNTER DB".Conveyor_C4_Collator.Maximum_Count;
      A     "B 6.7";
      =     #BIT0;
      A     "M 31.6";
      AN    "M 31.7";
      =     #XFER;
      CALL "DE-BOUNCER / COUNTER" (
           Bit_0                    := #BIT0,
           Bit_1                    := "B 7.0",
           Transfer_Start           := #XFER,
           Error_Reset              := "M 9.1",
           Space_DX_mS              := 600,
           ReSample_DX              := 85,
           Conveyor_Type            := 1,
           Preset_MIN_mS            := 500,
           LowSpd_Dimension_mS      := 0,
           HighSpd_Dimension_mS     := "HOUSE_KEEPING DB".C4_Packet_Length_mS,
           Plc_Scan_mS              := "DB UTILITY".Scan_Cycle_Previous,
           Q_Error                  := #ERROR,
           Word_Count               := "HMI_DB".CONV_4_COUNT,
           IO_DB                    := "DEBOUNCER COUNTER DB".Conveyor_C4_Collator);
M443: NOP   0;
NETWORK
TITLE =Packet Counter - Link Conveyor 5

      A     "A 45.0";
      L     S5T#1S;
      SF    "Timer 120"; // Call Hold 1s
      A     "Timer 120";
      =     "M 143.0";
      JNB   M450;
      L     "HMI_DB".CONVEYOR_MAXCOUNT_L;
      T     "DEBOUNCER COUNTER DB".Conveyor_C5_Link.Maximum_Count;
      A     "B 7.0";
      A     "M 35.1";
      AN    "M 35.2";
      =     #BIT0;
      A     "M 35.3";
      AN    "M 35.4";
      =     #XFER;
      CALL "DE-BOUNCER / COUNTER" (
           Bit_0                    := #BIT0,
           Bit_1                    := "B 7.1",
           Transfer_Start           := #XFER,
           Error_Reset              := "M 9.1",
           Space_DX_mS              := 600,
           ReSample_DX              := 85,
           Conveyor_Type            := 3,
           Preset_MIN_mS            := 500,
           LowSpd_Dimension_mS      := 0,
           HighSpd_Dimension_mS     := "HOUSE_KEEPING DB".C4_Packet_Length_mS,
           Plc_Scan_mS              := "DB UTILITY".Scan_Cycle_Previous,
           Q_Error                  := #ERROR,
           Word_Count               := "HMI_DB".CONV_5_COUNT,
           IO_DB                    := "DEBOUNCER COUNTER DB".Conveyor_C5_Link);
M450: NOP   0;
NETWORK
TITLE =Packet Counter - Delivery Conveyor 6

      A     "A 45.3";
      L     S5T#1S;
      SF    "Timer 121"; // Call Hold 1s
      A     "Timer 121";
      =     "M 143.1";
      JNB   M453;
      L     "HMI_DB".CONVEYOR_MAXCOUNT_L;
      T     "DEBOUNCER COUNTER DB".Conveyor_C6_Delivery.Maximum_Count;
      A     "B 7.1";
      A     "M 39.1";
      AN    "M 39.2";
      =     #BIT0;
      A     "M 39.4";
      AN    "M 39.5";
      =     #XFER;
      CALL "DE-BOUNCER / COUNTER" (
           Bit_0                    := #BIT0,
           Bit_1                    := "B 7.3",
           Transfer_Start           := #XFER,
           Error_Reset              := "M 9.1",
           Space_DX_mS              := 600,
           ReSample_DX              := 85,
           Conveyor_Type            := 2,
           Preset_MIN_mS            := 500,
           LowSpd_Dimension_mS      := 0,
           HighSpd_Dimension_mS     := "HOUSE_KEEPING DB".C4_Packet_Length_mS,
           Plc_Scan_mS              := "DB UTILITY".Scan_Cycle_Previous,
           Q_Error                  := #ERROR,
           Word_Count               := "HMI_DB".CONV_6_COUNT,
           IO_DB                    := "DEBOUNCER COUNTER DB".Conveyor_C6_Delivery);
M453: NOP   0;
NETWORK
TITLE =Packet Presence - Flipper / TurnTable / Conveyor 9 / Pusher 2

      L     0;
      A     "M 43.4";
      JCN   M434;
      L     1;
M434: T     "HMI_DB".FLIPPER_PACK_PRESENCE;
      T     "HMI_DB".FLIPPER_PACK_PRESENCE;
      L     0;
      A     "M 47.4";
      JCN   M474;
      L     1;
M474: T     "HMI_DB".TURNTABLE_PACK_PRESENCE;
      T     "HMI_DB".TURNTABLE_PACK_PRESENCE;
      L     0;
      A     "M 51.4";
      JCN   M514;
      L     1;
M514: T     "HMI_DB".ROLLER_PACK_PRESENCE;
      T     "HMI_DB".ROLLER_PACK_PRESENCE;
      L     0;
      A     "M 51.5";
      JCN   M515;
      L     1;
M515: T     "HMI_DB".PUSHER_PACK_PRESENCE;
      T     "HMI_DB".PUSHER_PACK_PRESENCE;
NETWORK
TITLE =Packet Counter - Pivot Conveyor 10

      A     "A 48.0";
      L     S5T#1S;
      SF    T    134; // Call Hold 1s
      A     T    134;
      JNB   M480;
      L     "HMI_DB".CONVEYOR_MAXCOUNT_W;
      T     "DEBOUNCER COUNTER DB".Conveyor_C10_Collator.Maximum_Count;
      A     "B 10.4";
      =     #BIT0;
      A     "M 55.5";
      AN    "M 55.6";
      =     #XFER;
      CALL "DE-BOUNCER / COUNTER" (
           Bit_0                    := #BIT0,
           Bit_1                    := "B 10.6",
           Transfer_Start           := #XFER,
           Error_Reset              := "M 9.1",
           Space_DX_mS              := 600,
           ReSample_DX              := 85,
           Conveyor_Type            := 1,
           Preset_MIN_mS            := 500,
           LowSpd_Dimension_mS      := 0,
           HighSpd_Dimension_mS     := #DIM_31,
           Plc_Scan_mS              := "DB UTILITY".Scan_Cycle_Previous,
           Q_Error                  := #ERROR,
           Word_Count               := "HMI_DB".CONV_10_COUNT,
           IO_DB                    := "DEBOUNCER COUNTER DB".Conveyor_C10_Collator);
M480: NOP   0;
NETWORK
TITLE =Packet Counter - Link Conveyor 11 (Low)

      A     "A 48.3";
      L     S5T#1S;
      SF    "Timer 122"; // Call Hold 1s
      A     "Timer 122";
      =     "M 143.2";
      JNB   M483;
      L     "HMI_DB".CONVEYOR_MAXCOUNT_W;
      T     "DEBOUNCER COUNTER DB".Conveyor_C11_Link.Maximum_Count;
      A     "B 10.6";
      A     "M 59.1";
      AN    "M 59.2";
      A     "P 15.1";
      =     #BIT0;
      A     "M 59.3";
      AN    "M 59.4";
      =     #XFER;
      CALL "DE-BOUNCER / COUNTER" (
           Bit_0                    := #BIT0,
           Bit_1                    := "B 10.7",
           Transfer_Start           := #XFER,
           Error_Reset              := "M 9.1",
           Space_DX_mS              := 600,
           ReSample_DX              := 85,
           Conveyor_Type            := 3,
           Preset_MIN_mS            := 300,
           LowSpd_Dimension_mS      := 0,
           HighSpd_Dimension_mS     := #DIM_31,
           Plc_Scan_mS              := "DB UTILITY".Scan_Cycle_Previous,
           Q_Error                  := #ERROR,
           Word_Count               := "HMI_DB".CONV_11_COUNT,
           IO_DB                    := "DEBOUNCER COUNTER DB".Conveyor_C11_Link);
M483: NOP   0;
NETWORK
TITLE =Packet Counter - Link Conveyor 12 (Low)

      A     "A 48.6";
      L     S5T#1S;
      SF    "Timer 123"; // Call Hold 1s
      A     "Timer 123";
      =     "M 143.3";
      JNB   M486;
      L     "HMI_DB".CONVEYOR_MAXCOUNT_W;
      T     "DEBOUNCER COUNTER DB".Conveyor_C12_Link.Maximum_Count;
      A     "B 10.7";
      A     "M 63.1";
      AN    "M 63.2";
      =     #BIT0;
      A     "M 63.3";
      AN    "M 63.4";
      =     #XFER;
      CALL "DE-BOUNCER / COUNTER" (
           Bit_0                    := #BIT0,
           Bit_1                    := "B 11.0",
           Transfer_Start           := #XFER,
           Error_Reset              := "M 9.1",
           Space_DX_mS              := 600,
           ReSample_DX              := 85,
           Conveyor_Type            := 3,
           Preset_MIN_mS            := 300,
           LowSpd_Dimension_mS      := 0,
           HighSpd_Dimension_mS     := #DIM_31,
           Plc_Scan_mS              := "DB UTILITY".Scan_Cycle_Previous,
           Q_Error                  := #ERROR,
           Word_Count               := "HMI_DB".CONV_12_COUNT,
           IO_DB                    := "DEBOUNCER COUNTER DB".Conveyor_C12_Link);
M486: NOP   0;
NETWORK
TITLE =Packet Counter - Delivery Conveyor 13 (Low)

      A     "A 49.0";
      L     S5T#1S;
      SF    "Timer 124"; // Call Hold 1s
      A     "Timer 124";
      =     "M 143.4";
      JNB   M490;
      L     "HMI_DB".CONVEYOR_MAXCOUNT_W;
      T     "DEBOUNCER COUNTER DB".Conveyor_C13_Delivery.Maximum_Count;
      A     "B 11.0";
      A     "M 67.1";
      AN    "M 67.2";
      =     #BIT0;
      A     "M 67.4";
      AN    "M 67.5";
      =     #XFER;
      CALL "DE-BOUNCER / COUNTER" (
           Bit_0                    := #BIT0,
           Bit_1                    := "B 11.2",
           Transfer_Start           := #XFER,
           Error_Reset              := "M 9.1",
           Space_DX_mS              := 600,
           ReSample_DX              := 85,
           Conveyor_Type            := 2,
           Preset_MIN_mS            := 300,
           LowSpd_Dimension_mS      := 0,
           HighSpd_Dimension_mS     := #DIM_237,
           Plc_Scan_mS              := "DB UTILITY".Scan_Cycle_Previous,
           Q_Error                  := #ERROR,
           Word_Count               := "HMI_DB".CONV_13_COUNT,
           IO_DB                    := "DEBOUNCER COUNTER DB".Conveyor_C13_Delivery);
M490: NOP   0;
NETWORK
TITLE =Packet Counter - Link Conveyor 21 (High)

      A     "A 53.4";
      L     S5T#1S;
      SF    "Timer 125"; // Call Hold 1s
      A     "Timer 125";
      =     "M 143.5";
      JNB   M534;
      L     "HMI_DB".CONVEYOR_MAXCOUNT_W;
      T     "DEBOUNCER COUNTER DB".Conveyor_C21_Link.Maximum_Count;
      A     "B 10.6";
      A     "M 79.1";
      AN    "M 79.2";
      A     "P 15.0";
      =     #BIT0;
      A     "M 79.3";
      AN    "M 79.4";
      =     #XFER;
      CALL "DE-BOUNCER / COUNTER" (
           Bit_0                    := #BIT0,
           Bit_1                    := "B 15.4",
           Transfer_Start           := #XFER,
           Error_Reset              := "M 9.1",
           Space_DX_mS              := 600,
           ReSample_DX              := 85,
           Conveyor_Type            := 3,
           Preset_MIN_mS            := 300,
           LowSpd_Dimension_mS      := 0,
           HighSpd_Dimension_mS     := #DIM_31,
           Plc_Scan_mS              := "DB UTILITY".Scan_Cycle_Previous,
           Q_Error                  := #ERROR,
           Word_Count               := "HMI_DB".CONV_21_COUNT,
           IO_DB                    := "DEBOUNCER COUNTER DB".Conveyor_C21_Link);
M534: NOP   0;
NETWORK
TITLE =Packet Counter - Link Conveyor 22 (High)

      A     "A 53.6";
      L     S5T#1S;
      SF    "Timer 126"; // Call Hold 1s
      A     "Timer 126";
      =     "M 143.6";
      JNB   M536;
      L     "HMI_DB".CONVEYOR_MAXCOUNT_W;
      T     "DEBOUNCER COUNTER DB".Conveyor_C22_Link.Maximum_Count;
      A     "B 15.4";
      A     "M 83.1";
      AN    "M 83.2";
      =     #BIT0;
      A     "M 83.3";
      AN    "M 83.4";
      =     #XFER;
      CALL "DE-BOUNCER / COUNTER" (
           Bit_0                    := #BIT0,
           Bit_1                    := "B 15.5",
           Transfer_Start           := #XFER,
           Error_Reset              := "M 9.1",
           Space_DX_mS              := 600,
           ReSample_DX              := 85,
           Conveyor_Type            := 3,
           Preset_MIN_mS            := 300,
           LowSpd_Dimension_mS      := 0,
           HighSpd_Dimension_mS     := #DIM_31,
           Plc_Scan_mS              := "DB UTILITY".Scan_Cycle_Previous,
           Q_Error                  := #ERROR,
           Word_Count               := "HMI_DB".CONV_22_COUNT,
           IO_DB                    := "DEBOUNCER COUNTER DB".Conveyor_C22_Link);
M536: NOP   0;
NETWORK
TITLE =Packet Counter - Delivery Conveyor 23 (High)

      A     "A 54.0";
      L     S5T#1S;
      SF    "Timer 127"; // Call Hold 1s
      A     "Timer 127";
      =     "M 143.7";
      JNB   M540;
      L     "HMI_DB".CONVEYOR_MAXCOUNT_W;
      T     "DEBOUNCER COUNTER DB".Conveyor_C23_Delivery.Maximum_Count;
      A     "B 15.5";
      A     "M 87.1";
      AN    "M 87.2";
      =     #BIT0;
      A     "M 87.4";
      AN    "M 87.5";
      =     #XFER;
      CALL "DE-BOUNCER / COUNTER" (
           Bit_0                    := #BIT0,
           Bit_1                    := "B 15.7",
           Transfer_Start           := #XFER,
           Error_Reset              := "M 9.1",
           Space_DX_mS              := 600,
           ReSample_DX              := 85,
           Conveyor_Type            := 2,
           Preset_MIN_mS            := 300,
           LowSpd_Dimension_mS      := 0,
           HighSpd_Dimension_mS     := #DIM_237,
           Plc_Scan_mS              := "DB UTILITY".Scan_Cycle_Previous,
           Q_Error                  := #ERROR,
           Word_Count               := "HMI_DB".CONV_23_COUNT,
           IO_DB                    := "DEBOUNCER COUNTER DB".Conveyor_C23_Delivery);
M540: NOP   0;
NETWORK
TITLE =HMI Packet Counters Reset (Same Conditions as FC1206)
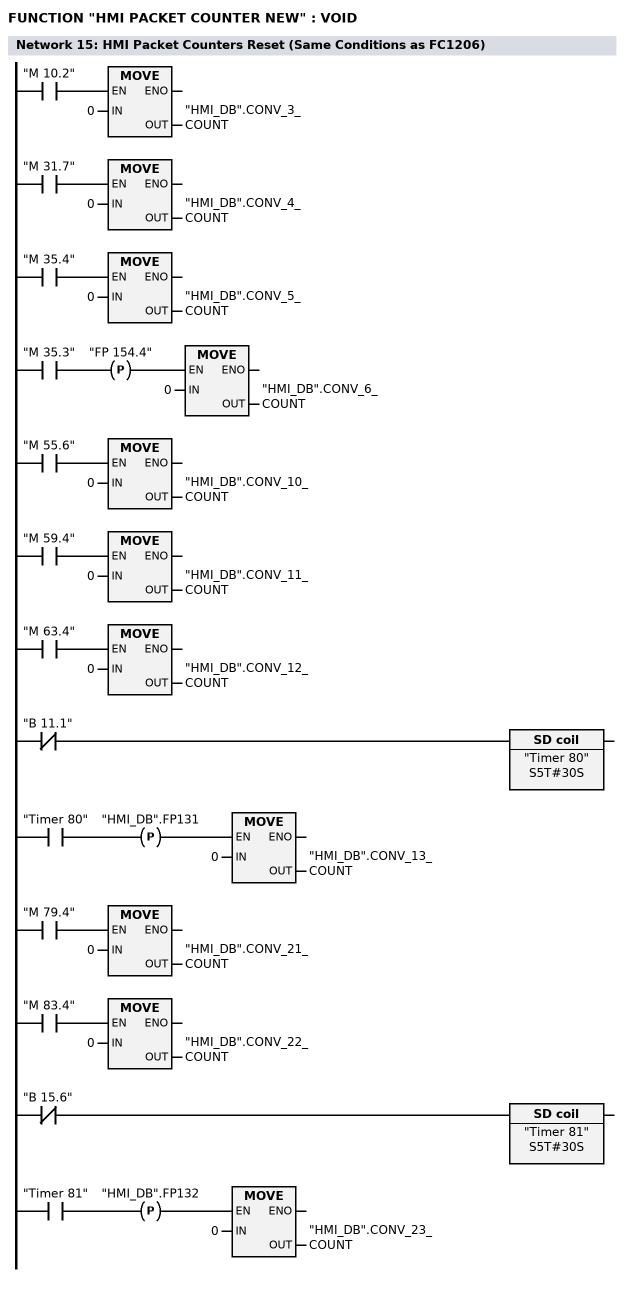

      A     "M 10.2";
      JNB   F102;
      L     0;
      T     "HMI_DB".CONV_3_COUNT; // FC8 Takes Over 0 on Next Call
F102: NOP   0;
      A     "M 31.7";
      JNB   F317;
      L     0;
      T     "HMI_DB".CONV_4_COUNT; // FC8 Takes Over 0 on Next Call
F317: NOP   0;
      A     "M 35.4";
      JNB   F354;
      L     0;
      T     "HMI_DB".CONV_5_COUNT; // FC8 Takes Over 0 on Next Call
F354: NOP   0;
      A     "M 35.3";
      FP    "FP 154.4";
      JNB   F396;
      L     0;
      T     "HMI_DB".CONV_6_COUNT; // FC8 Takes Over 0 on Next Call
F396: NOP   0;
      A     "M 55.6";
      JNB   F556;
      L     0;
      T     "HMI_DB".CONV_10_COUNT; // FC8 Takes Over 0 on Next Call
F556: NOP   0;
      A     "M 59.4";
      JNB   F594;
      L     0;
      T     "HMI_DB".CONV_11_COUNT; // FC8 Takes Over 0 on Next Call
F594: NOP   0;
      A     "M 63.4";
      JNB   F634;
      L     0;
      T     "HMI_DB".CONV_12_COUNT; // FC8 Takes Over 0 on Next Call
F634: NOP   0;
      AN    "B 11.1";
      L     S5T#30S;
      SD    "Timer 80";
      A     "Timer 80";
      FP    "HMI_DB".FP131;
      JNB   F676;
      L     0;
      T     "HMI_DB".CONV_13_COUNT; // FC8 Takes Over 0 on Next Call
F676: NOP   0;
      A     "M 79.4";
      JNB   F794;
      L     0;
      T     "HMI_DB".CONV_21_COUNT; // FC8 Takes Over 0 on Next Call
F794: NOP   0;
      A     "M 83.4";
      JNB   F834;
      L     0;
      T     "HMI_DB".CONV_22_COUNT; // FC8 Takes Over 0 on Next Call
F834: NOP   0;
      AN    "B 15.6";
      L     S5T#30S;
      SD    "Timer 81";
      A     "Timer 81";
      FP    "HMI_DB".FP132;
      JNB   F876;
      L     0;
      T     "HMI_DB".CONV_23_COUNT; // FC8 Takes Over 0 on Next Call
F876: NOP   0;
END_FUNCTION

FUNCTION "FM350 COUNTERS" : VOID
TITLE =Counters
//FM350-2 : Counter Module Added to measure Collator Conveyors 4 & 10 Filling
//Surface Left, and to measure Packets Length & Width in order to Fit the Most
//Packets Number onto the Respective Conveyor... May 22
VERSION : 0.1


VAR_TEMP
  ENCODER_STOP : BOOL ;
  RETURN_RD : INT ;	//Print Pulse Read Function Return
  PRESS_LENGTH_3 : WORD ;	//Slat Conveyor 3 - Surface per Packet
  PACKET_LENGTH_4 : WORD ;	//Collator Conveyor 4 - Packet Length
  HALF_PACKET_LENGTH_4 : WORD ;	//Collator Conveyor 4 - Packet Length - Half
  PACKET_LENGTH_HALF_4 : WORD ;	//Collator Conveyor 4 - Packet Length + Half
  SURFACE_LENGTH_LEFT_4 : WORD ;	//Collator Conveyor 4 - Surface Length Left
  QTY_MAX_4 : REAL ;
  PACKET_WIDTH_10 : WORD ;	//Collator Conveyor 10 - Packet Width
  HALF_PACKET_WIDTH_10 : WORD ;	//Collator Conveyor 10 - Packet Width - Half
  PACKET_WIDTH_HALF_10 : WORD ;	//Collator Conveyor 10 - Packet Width + Half
  SURFACE_LENGTH_LEFT_10 : WORD ;
  QTY_MAX_10 : WORD ;
END_VAR
BEGIN
NETWORK
TITLE =Call DB

      OPN   "FM350 DB";
      CALL "CNT2_CTR" (//Control the FM 350-2
           DB_NO                    := W#16#2);

NETWORK
TITLE =FM350-2 Address Resets

      A     "M 167.7";
      JNB   M677;
      L     W#16#140;
      T     DBW   12;
//;
      L     DW#16#A00;
      T     DBD   14;
//;
      R     "M 167.7";

M677: NOP   0;
NETWORK
TITLE =Read Counters Jobs
//FM350-2 :  Job 100 = Read Counter 0,1,2,3
//           Job 101 = Read Counter 4,5,6,7
//           Then Transfer to DB2
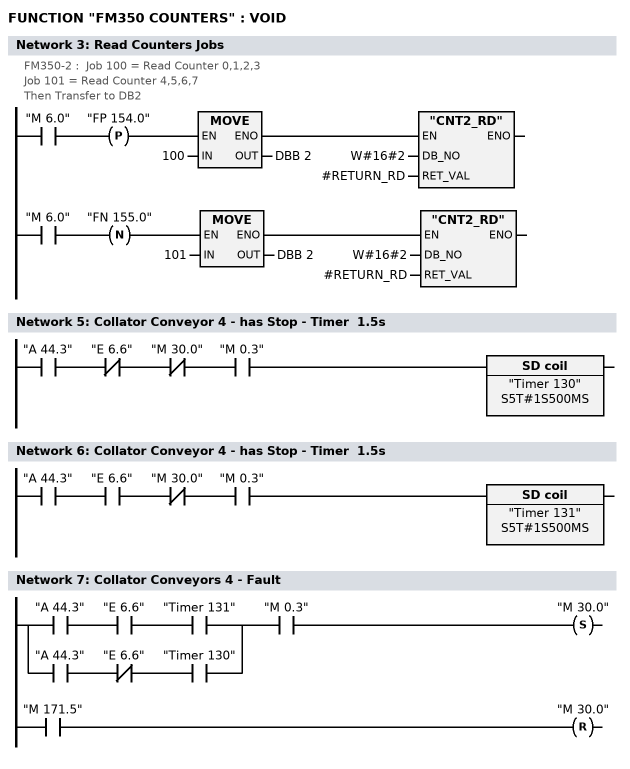
      A     "M 6.0";
      FP    "FP 154.0";
      JNB   M154;
      L     100;
      T     DBB    2;
      CALL "CNT2_RD" (
           DB_NO                    := W#16#2,
           RET_VAL                  := #RETURN_RD);

M154: NOP   0;

      A     "M 6.0";
      FN    "FN 155.0";
      JNB   M155;
      L     101;
      T     DBB    2;
      CALL "CNT2_RD" (
           DB_NO                    := W#16#2,
           RET_VAL                  := #RETURN_RD);

M155: NOP   0;
NETWORK
TITLE =
//Encoder Health Monitor


NETWORK
TITLE =Collator Conveyor 4 - has Stop - Timer  1.5s

      A     "A 44.3";
      AN    "E 6.6";
      AN    "M 30.0";
      A     "M 0.3";
      L     S5T#1S500MS;
      SD    "Timer 130";
NETWORK
TITLE =Collator Conveyor 4 - has Stop - Timer  1.5s

      A     "A 44.3";
      A     "E 6.6";
      AN    "M 30.0";
      A     "M 0.3";
      L     S5T#1S500MS;
      SD    "Timer 131";
NETWORK
TITLE =Collator Conveyors 4 - Fault

      A(    ;
      A     "A 44.3";
      A     "E 6.6";
      A     "Timer 131";
      O     ;
      A     "A 44.3";
      AN    "E 6.6";
      A     "Timer 130";
      )     ;
      A     "M 0.3";
      S     "M 30.0";
//;
      O     "M 171.5";
      R     "M 30.0";
NETWORK
TITLE =Collator Conveyors 4 - Lauer Comm

      OPN   "DB LAUER";

      A     "E 6.6";
      JC    M001;

      L     2#0;
      T     DBW  232;
      JU    M002;

M001: L     2#1;
      T     DBW  232;

M002: NOP   0;
END_FUNCTION

FUNCTION "ELEVATOR TEST FUNCTION" : VOID
TITLE =
VERSION : 0.1

BEGIN
NETWORK
TITLE =


      A     "A 63.0";
      JCN   M003;
      A     "A 63.3";
      JCN   M002;
      L     MW   950;
      L     1;
      -I    ;
      T     MW   950;
      JU    M001;
M002: L     MW   950;
      L     1;
      +I    ;
      T     MW   950;
M001: L     MW   950;
      L     200;
      <=I   ;
      =     M    930.1;
      L     MW   950;
      L     10;
      <=I   ;
      =     M    930.0;
      L     MW   950;
      L     800;
      >=I   ;
      =     M    930.2;
      L     MW   950;
      L     990;
      >=I   ;
      =     M    930.3;
M003: CLR   ;


END_FUNCTION

ORGANIZATION_BLOCK "CYCLIC"
TITLE =Main Cycle
VERSION : 0.0


VAR_TEMP
  OB1_EV_CLASS : BYTE ;	//Bits 0-3 = 1 (Coming event), Bits 4-7 = 1 (Event class 1)
  OB1_SCAN_1 : BYTE ;	//1 (Cold restart scan 1 of OB 1), 3 (Scan 2-n of OB 1)
  OB1_PRIORITY : BYTE ;	//1 (Priority of 1 is lowest)
  OB1_OB_NUMBR : BYTE ;	//1 (Organization block 1, OB1)
  OB1_RESERVED_1 : BYTE ;	//Reserved for system
  OB1_RESERVED_2 : BYTE ;	//Reserved for system
  OB1_PREV_CYCLE : INT ;	//Cycle time of previous OB1 scan (milliseconds)
  OB1_MIN_CYCLE : INT ;	//Minimum cycle time of OB1 (milliseconds)
  OB1_MAX_CYCLE : INT ;	//Maximum cycle time of OB1 (milliseconds)
  OB1_DATE_TIME : DATE_AND_TIME ;	//Date and time OB1 started
END_VAR
BEGIN
NETWORK
TITLE =Scan Time
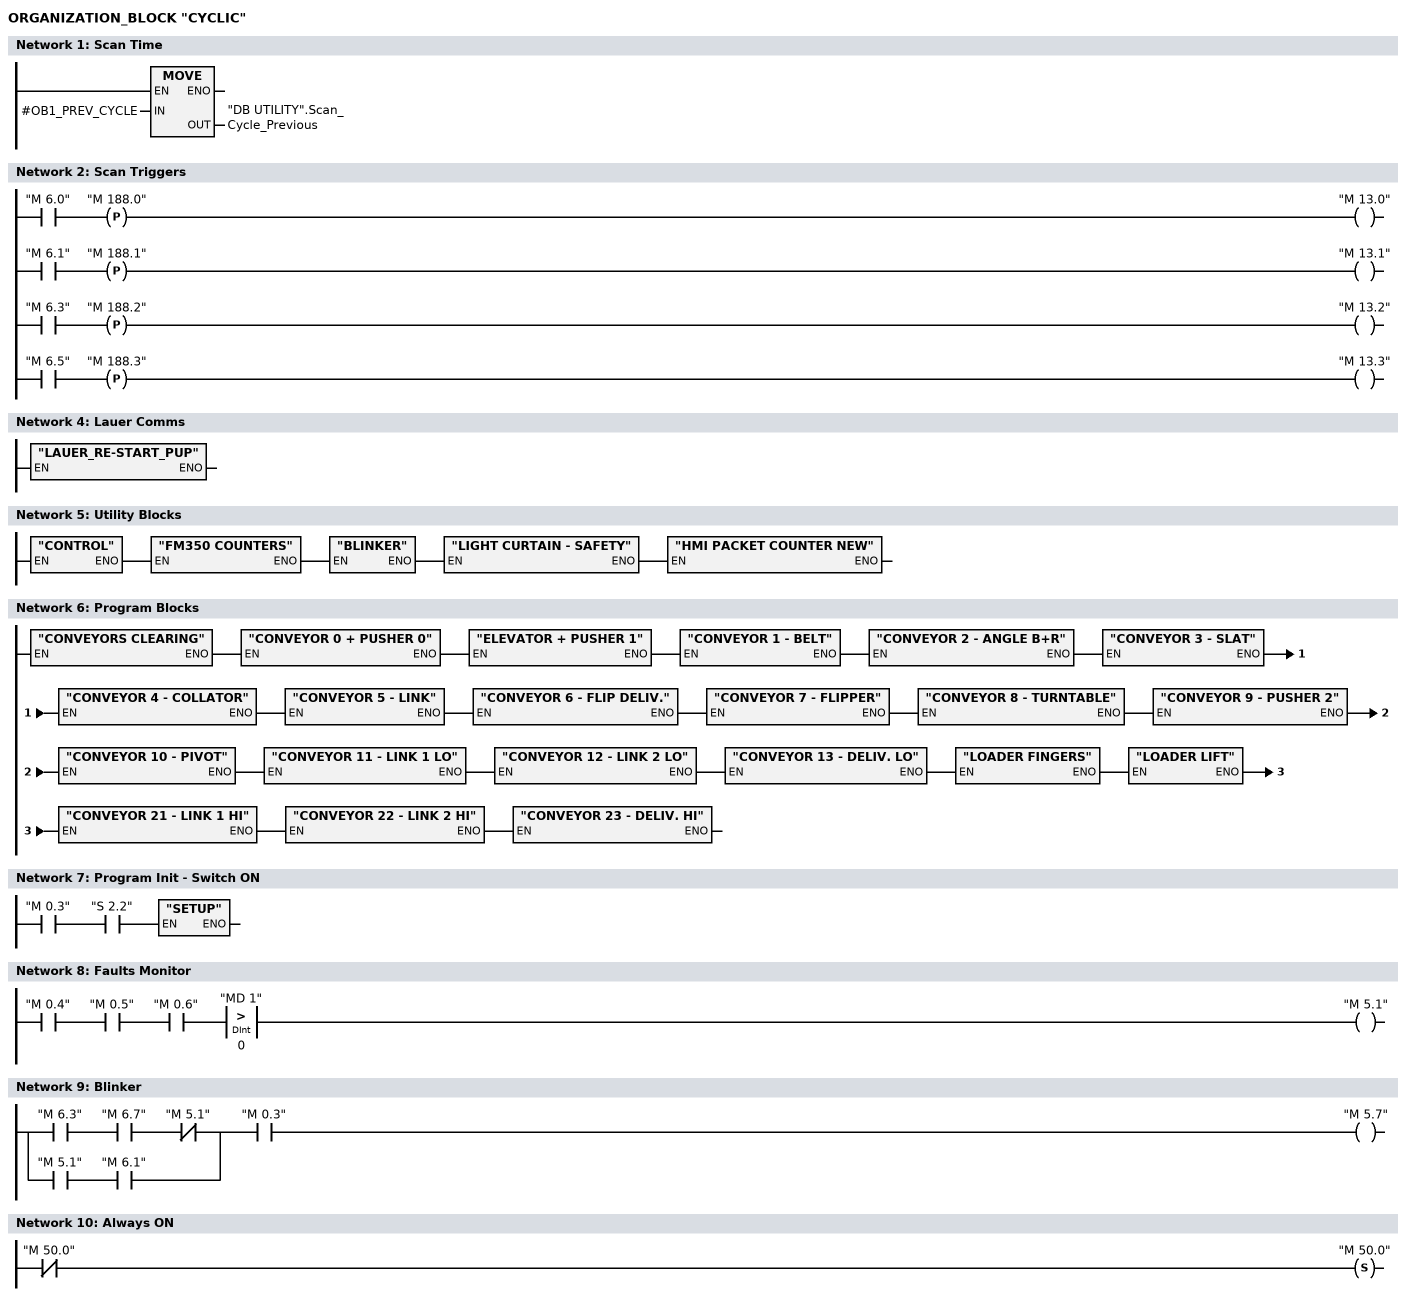

      L     #OB1_PREV_CYCLE;
      T     "DB UTILITY".Scan_Cycle_Previous;
NETWORK
TITLE =Scan Triggers

      A     "M 6.0";
      FP    "M 188.0";
      =     "M 13.0";
//;
      A     "M 6.1";
      FP    "M 188.1";
      =     "M 13.1";
//;
      A     "M 6.3";
      FP    "M 188.2";
      =     "M 13.2";
//;
      A     "M 6.5";
      FP    "M 188.3";
      =     "M 13.3";
NETWORK
TITLE =Packet Counters
//     CALL  "HMI PACKET COUNTER OLD"



//  CALL  "ELEVATOR TEST FUNCTION"

NETWORK
TITLE =Lauer Comms

      CALL "LAUER_RE-START_PUP" ;

NETWORK
TITLE =Utility Blocks

      CALL "CONTROL" ;
      CALL "FM350 COUNTERS" ;
      CALL "BLINKER" ;
      CALL "LIGHT CURTAIN - SAFETY" ;
      CALL "HMI PACKET COUNTER  NEW" ;
NETWORK
TITLE =Program Blocks

      CALL "CONVEYORS CLEARING" ;

      CALL "CONVEYOR 0 + PUSHER 0" ;
      CALL "ELEVATOR + PUSHER 1" ;
      CALL "CONVEYOR 1 - BELT" ;
      CALL "CONVEYOR 2 - ANGLE B+R" ;
      CALL "CONVEYOR 3 - SLAT" ;
      CALL "CONVEYOR 4 - COLLATOR" ;
      CALL "CONVEYOR 5 - LINK" ;

      CALL "CONVEYOR 6 - FLIP DELIV." ;
      CALL "CONVEYOR 7 - FLIPPER" ;

      CALL "CONVEYOR 8 - TURNTABLE" ;

      CALL "CONVEYOR 9 - PUSHER 2" ;
      CALL "CONVEYOR 10 - PIVOT" ;
      CALL "CONVEYOR 11 - LINK 1 LO" ;
      CALL "CONVEYOR 12 - LINK 2 LO" ;
      CALL "CONVEYOR 13 - DELIV. LO" ;
      CALL "LOADER FINGERS" ;
      CALL "LOADER LIFT" ;
      CALL "CONVEYOR 21 - LINK 1 HI" ;
      CALL "CONVEYOR 22 - LINK 2 HI" ;
      CALL "CONVEYOR 23 - DELIV. HI" ;


NETWORK
TITLE =Program Init - Switch ON

      A     "M 0.3";
      A     "S 2.2";
      JNB   M022;
      CALL "SETUP" ;

M022: NOP   0;
NETWORK
TITLE =Faults Monitor

      A     "M 0.4";
      A     "M 0.5";
      A     "M 0.6";
      A(    ;
      L     "MD 1";
      L     0;
      >D    ;
      )     ;
      =     "M 5.1";
NETWORK
TITLE =Blinker

      A(    ;
      A     "M 6.3";
      A     "M 6.7";
      AN    "M 5.1";
      O     ;
      A     "M 5.1";
      A     "M 6.1";
      )     ;
      A     "M 0.3";
      =     "M 5.7";
NETWORK
TITLE =Always ON

      AN    "M 50.0";
      S     "M 50.0";
END_ORGANIZATION_BLOCK

ORGANIZATION_BLOCK "Cyclic 100mS"
TITLE = "Cyclic Interrupt"
VERSION : 0.1


VAR_TEMP
  OB35_EV_CLASS : BYTE ;	//Bits 0-3 = 1 (Coming event), Bits 4-7 = 1 (Event class 1)
  OB35_STRT_INF : BYTE ;	//16#36 (OB 35 has started)
  OB35_PRIORITY : BYTE ;	//Priority of OB Execution
  OB35_OB_NUMBR : BYTE ;	//35 (Organization block 35, OB35)
  OB35_RESERVED_1 : BYTE ;	//Reserved for system
  OB35_RESERVED_2 : BYTE ;	//Reserved for system
  OB35_PHASE_OFFSET : WORD ;	//Phase offset (msec)
  OB35_RESERVED_3 : INT ;	//Reserved for system
  OB35_EXC_FREQ : INT ;	//Frequency of execution (msec)
  OB35_DATE_TIME : DATE_AND_TIME ;	//Date and time OB35 started
END_VAR
BEGIN
NETWORK
TITLE =CYCLIC 100 mS

      CALL "GENERAL FAULTS" ;
      CALL "HMI CONTROL" ;
      CALL "HMI COMMS" ;
      CALL "LIGHT BAR" ;

//  CALL  "Sensor Check Calls"
NETWORK
TITLE =Lauer Comms

      CALL "LAUER CALL" ;

NETWORK
TITLE =Lauer Comms

      CALL "LAUER COMM FC" (
           UBDB                     := "DB LAUER",
           RXFA                     := 36,
           RXLE                     := 32,
           TXFA                     := 3,
           TXLE                     := 32,
           RSET                     := "M 210.1",
           TIMT                     := T    105,
           TIMZ                     := S5T#1S,
           COFF                     := "LAUER RESTART FC",
           INIT                     := "LAUER COMM ERR FC",
           RFLM                     := "M 210.0",
           EROR                     := "M 210.2");
END_ORGANIZATION_BLOCK

ORGANIZATION_BLOCK "I/O_FLT1"
TITLE = "I/O Point Fault"
VERSION : 0.1


VAR_TEMP
  OB82_EV_CLASS : BYTE ;	//16#39, Event class 3, Entering event state, Internal fault event
  OB82_FLT_ID : BYTE ;	//16#XX, Fault identifcation code
  OB82_PRIORITY : BYTE ;	//Priority of OB Execution
  OB82_OB_NUMBR : BYTE ;	//82 (Organization block 82, OB82)
  OB82_RESERVED_1 : BYTE ;	//Reserved for system
  OB82_IO_FLAG : BYTE ;	//Input (01010100), Output (01010101)
  OB82_MDL_ADDR : WORD ;	//Base address of module with fault
  OB82_MDL_DEFECT : BOOL ;	//Module defective
  OB82_INT_FAULT : BOOL ;	//Internal fault
  OB82_EXT_FAULT : BOOL ;	//External fault
  OB82_PNT_INFO : BOOL ;	//Point information
  OB82_EXT_VOLTAGE : BOOL ;	//External voltage low
  OB82_FLD_CONNCTR : BOOL ;	//Field wiring connector missing
  OB82_NO_CONFIG : BOOL ;	//Module has no configuration data
  OB82_CONFIG_ERR : BOOL ;	//Module has configuration error
  OB82_MDL_TYPE : BYTE ;	//Type of module
  OB82_SUB_MDL_ERR : BOOL ;	//Sub-Module is missing or has error
  OB82_COMM_FAULT : BOOL ;	//Communication fault
  OB82_MDL_STOP : BOOL ;	//Module is stopped
  OB82_WTCH_DOG_FLT : BOOL ;	//Watch dog timer stopped module
  OB82_INT_PS_FLT : BOOL ;	//Internal power supply fault
  OB82_PRIM_BATT_FLT : BOOL ;	//Primary battery is in fault
  OB82_BCKUP_BATT_FLT : BOOL ;	//Backup battery is in fault
  OB82_RESERVED_2 : BOOL ;	//Reserved for system
  OB82_RACK_FLT : BOOL ;	//Rack fault, only for bus interface module
  OB82_PROC_FLT : BOOL ;	//Processor fault
  OB82_EPROM_FLT : BOOL ;	//EPROM fault
  OB82_RAM_FLT : BOOL ;	//RAM fault
  OB82_ADU_FLT : BOOL ;	//ADU fault
  OB82_FUSE_FLT : BOOL ;	//Fuse fault
  OB82_HW_INTR_FLT : BOOL ;	//Hardware interupt input in fault
  OB82_RESERVED_3 : BOOL ;	//Reserved for system
  OB82_DATE_TIME : DATE_AND_TIME ;	//Date and time OB82 started
END_VAR
BEGIN
NETWORK
TITLE =

END_ORGANIZATION_BLOCK

ORGANIZATION_BLOCK "RACK_FLT"
TITLE = "Loss Of Rack Fault"
VERSION : 0.1


VAR_TEMP
  OB86_EV_CLASS : BYTE ;	//16#38/39 Event class 3
  OB86_FLT_ID : BYTE ;	//16#C1/C4/C5, Fault identifcation code
  OB86_PRIORITY : BYTE ;	//Priority of OB Execution
  OB86_OB_NUMBR : BYTE ;	//86 (Organization block 86, OB86)
  OB86_RESERVED_1 : BYTE ;	//Reserved for system
  OB86_RESERVED_2 : BYTE ;	//Reserved for system
  OB86_MDL_ADDR : WORD ;	//Base address of IM module in rack with fault
  OB86_RACKS_FLTD : ARRAY  [0 .. 31 ] OF BOOL ;	//Racks in fault
  OB86_DATE_TIME : DATE_AND_TIME ;	//Date and time OB86 started
END_VAR
BEGIN
NETWORK
TITLE =

END_ORGANIZATION_BLOCK

ORGANIZATION_BLOCK "OB100"
TITLE =Start up    OB100
VERSION : 0.1


VAR_TEMP
  OB100_EV_CLASS : BYTE ;	//16#13, Event class 1, Entering event state, Event logged in diagnostic buffer
  OB100_STRTUP : BYTE ;	//16#81/82/83/84 Method of startup
  OB100_PRIORITY : BYTE ;	//27 (Priority of 1 is lowest)
  OB100_OB_NUMBR : BYTE ;	//100 (Organization block 100, OB100)
  OB100_RESERVED_1 : BYTE ;	//Reserved for system
  OB100_RESERVED_2 : BYTE ;	//Reserved for system
  OB100_STOP : WORD ;	//Event that caused CPU to stop (16#4xxx)
  OB100_STRT_INFO : DWORD ;	//Information on how system started
  OB100_DATE_TIME : DATE_AND_TIME ;	//Date and time OB100 started
END_VAR
BEGIN
NETWORK
TITLE =Lauer restart bit

      L     2#0; // Reset First cycle Flag
      =     "M 210.0";
NETWORK
TITLE =HMI On Lamp

      AN    "HMI_DB".AERIAL_LINK_RUN_PB;
      =     "HMI_DB".AERIAL_LINK_RUN_PB;
NETWORK
TITLE =DB Init

      R     "DEBOUNCER COUNTER DB".Conveyor_C3_Slat.FirstScan_Done;
      R     "DEBOUNCER COUNTER DB".Conveyor_C4_Collator.FirstScan_Done;
      R     "DEBOUNCER COUNTER DB".Conveyor_C5_Link.FirstScan_Done;
      R     "DEBOUNCER COUNTER DB".Conveyor_C6_Delivery.FirstScan_Done;
      R     "DEBOUNCER COUNTER DB".Conveyor_C10_Collator.FirstScan_Done;
      R     "DEBOUNCER COUNTER DB".Conveyor_C11_Link.FirstScan_Done;
      R     "DEBOUNCER COUNTER DB".Conveyor_C12_Link.FirstScan_Done;
      R     "DEBOUNCER COUNTER DB".Conveyor_C13_Delivery.FirstScan_Done;
      R     "DEBOUNCER COUNTER DB".Conveyor_C21_Link.FirstScan_Done;
      R     "DEBOUNCER COUNTER DB".Conveyor_C22_Link.FirstScan_Done;
      R     "DEBOUNCER COUNTER DB".Conveyor_C23_Delivery.FirstScan_Done;
END_ORGANIZATION_BLOCK

ORGANIZATION_BLOCK "PROG_ERR"
TITLE = "Programming Error"
VERSION : 0.1


VAR_TEMP
  OB121_EV_CLASS : BYTE ;	//16#25, Event class 2, Entering event state, Internal fault event
  OB121_SW_FLT : BYTE ;	//16#XX Software programming fault
  OB121_PRIORITY : BYTE ;	//Priority of OB Execution
  OB121_OB_NUMBR : BYTE ;	//121 (Organization block 121, OB121)
  OB121_BLK_TYPE : BYTE ;	//16#88/8A/8B/8C/8E Type of block fault occured in
  OB121_RESERVED_1 : BYTE ;	//Reserved for system
  OB121_FLT_REG : WORD ;	//16#XX Specific register that caused fault
  OB121_BLK_NUM : WORD ;	//Number of block that programming fault occured in
  OB121_PRG_ADDR : WORD ;	//Address in block where programming fault occured
  OB121_DATE_TIME : DATE_AND_TIME ;	//Date and time OB121 started
END_VAR
BEGIN
NETWORK
TITLE =

END_ORGANIZATION_BLOCK

ORGANIZATION_BLOCK "IO ACCESS_ERR"
TITLE = "Programming Error"
VERSION : 0.1


VAR_TEMP
  OB121_EV_CLASS : BYTE ;	//16#25, Event class 2, Entering event state, Internal fault event
  OB121_SW_FLT : BYTE ;	//16#XX Software programming fault
  OB121_PRIORITY : BYTE ;	//Priority of OB Execution
  OB121_OB_NUMBR : BYTE ;	//121 (Organization block 121, OB121)
  OB121_BLK_TYPE : BYTE ;	//16#88/8A/8B/8C/8E Type of block fault occured in
  OB121_RESERVED_1 : BYTE ;	//Reserved for system
  OB121_FLT_REG : WORD ;	//16#XX Specific register that caused fault
  OB121_BLK_NUM : WORD ;	//Number of block that programming fault occured in
  OB121_PRG_ADDR : WORD ;	//Address in block where programming fault occured
  OB121_DATE_TIME : DATE_AND_TIME ;	//Date and time OB121 started
END_VAR
BEGIN
NETWORK
TITLE =

END_ORGANIZATION_BLOCK

